Fanuc KAREL source: kt00718.KL

-- PROVISIONAL review KL for V770-1; original PC SHA256 99aa0181adf50b620af600d2a11eb6e2823b2f9709162105b8469e777794f979
-- Incomplete behavior may be omitted. Consult companion uncertainty JSON. Do not deploy.
PROGRAM KT00718
%NOLOCKGROUP
VAR
  OUT : BOOLEAN
-- UNRESOLVED_DECL P1 type=000101
-- UNRESOLVED_DECL P2 type=000101
BEGIN
  -- UNRESOLVED_PC offsets 5-20; opcodes 22,63,23
  -- UNRESOLVED_PC offsets 25-29; opcodes 7F
END KT00718
